ABB RAPID module: MainCall.mod

%%%
  VERSION:1
  LANGUAGE:ENGLISH
%%%
MODULE MOD_MainCall

    ! -------------------------------
    ! Define customized variables here
    ! ...

	! Tool variables:

	! Reference variables:
	PERS wobjdata FrameS := [FALSE, TRUE, "", [[0,0,0],[1,0,0,0]],[[1234.570,-98.765,50.500],[0.96592583,0.00000000,0.00000000,0.25881905]]];

	PROC SubProg2()
		ConfJ \On;
		ConfL \Off;
		MoveAbsJ [[30.000000,25.000000,80.000000,-45.000000,0.000000,0.000000],[9E+09,9E+09,9E+09,9E+09,9E+09,9E+09]],v500,z1,tool0 \WObj:=FrameS;
	ENDPROC

	PROC Main()
		ConfJ \On;
		ConfL \Off;
		! Program generated by RoboDK v6.0.7 for ABB IRB 260 on XX/XX/XXXX 18:00:00
		! Using nominal kinematics.
		MoveAbsJ [[10.000000,-20.000000,50.000000,30.000000,0.000000,0.000000],[9E+09,9E+09,9E+09,9E+09,9E+09,9E+09]],v500,z1,tool0 \WObj:=FrameS;
		SubProg2;
		NotAProgram;
	ENDPROC

ENDMODULE
